Fanuc KAREL source: KT00479.KL

PROGRAM KT00479
%NOLOCKGROUP
VAR
  P1: POSITION
  P2: XYZWPR
  OUT: POSITION
BEGIN
    P2.Y = 2.0
  OUT = P1 : P2
END KT00479
